FUNCTION_BLOCK FsInfo (* Query the properties of the file server and the status of a volume *)
  (* Standard: 61499-2; Description: Uses iso_FscGetServerProperties(), iso_FscGetVolumeStatus() and iso_FscGetCurrentDirectory() of the CCI ISOBUS driver (ISO 11783-13). \n The space is the one of the volume of the current directory. u8VolumeStatus is 255 if the server has no volume status (e.g. version 3). \n Client is NmDestin.s16OwnCfHnd, file server is NmDestin.s16Handle (e.g. found with NmGetCfInfo, NAME function 61). \n The FB opens its own io channel to the server and closes it at the end. One job at a time: REQ during a job gives ERR with s16Status E_BUSY. \n Every REQ ends with exactly one CNF or ERR. *)
  (* Version 1.0, 2026-11-26, Franz Höpfinger, initial API and implementation and/or initial documentation *)
  PACKAGE isobus::fs;
  IMPORT isobus::pgn::ISONETEVENT_T;
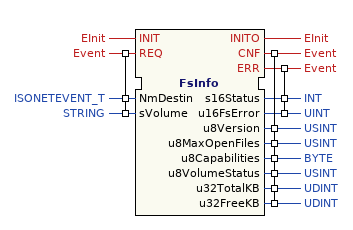
  EVENT_INPUT
    INIT : EInit; (* Service Initialization *)
    REQ WITH NmDestin, sVolume; (* Query the file server *)
  END_EVENT
  EVENT_OUTPUT
    INITO : EInit; (* Initialization Confirm *)
    CNF WITH u8Version, u8MaxOpenFiles, u8Capabilities, u8VolumeStatus, u32TotalKB, u32FreeKB; (* Properties read *)
    ERR WITH s16Status, u16FsError; (* Job failed *)
  END_EVENT
  VAR_INPUT
    NmDestin : isobus::pgn::ISONETEVENT_T; (* Client (s16OwnCfHnd) and file server (s16Handle) *)
    sVolume : STRING; (* Volume for the volume status, e.g. \\USB\, empty = volume of the current directory *)
  END_VAR
  VAR_OUTPUT
    s16Status : INT; (* With ERR: driver return value or own error (E_BUSY, E_RANGE, E_CONFIG) *)
    u16FsError : UINT; (* With ERR: file server or client error (ISO 11783-13 B.9, 6400 ff. client) *)
    u8Version : USINT; (* Version of the file server (3 = second edition, 4 = 2022) *)
    u8MaxOpenFiles : USINT; (* Maximum number of open files *)
    u8Capabilities : BYTE; (* Capabilities (ISO 11783-13 B.7) *)
    u8VolumeStatus : USINT; (* 0 present, 1 in use, 2 prepared for removal, 3 removed, 255 unknown *)
    u32TotalKB : UDINT; (* Size of the volume in KB *)
    u32FreeKB : UDINT; (* Free space of the volume in KB *)
  END_VAR
END_FUNCTION_BLOCK
